# EPICS SNL sequencer program: injectorApp/src/injectorRampe_C2.stt
/*
#  C.E.A. IRFU/SIS/LDISC
#
#
#
*/
/*
*-----------------------------------------------------------------------
*   IFMIF/EVEDA Injecteur:
*   snl_Rampe_C2 : programme SNL pour la gestion de la commande de
*            rampe de COIL02_PS
*-----------------------------------------------------------------------
*/

/*program snl_Rampe_C2*/

program injectorRampe_C2

short OK_Rampe;
assign OK_Rampe to "SRC:COIL02_PS:PretRampe";
monitor OK_Rampe;

short Envoi_Rampe;
assign Envoi_Rampe to "SRC:COIL02_PS:RampeCmd";
monitor Envoi_Rampe;

ss ss1
{

        state connected {
             when ( (delay(2.0)) && (pvConnectCount() == pvChannelCount()) ) {
              printf("SNL_Rampe_C2 :entree programme - connexions etablies \n");

             } state Debut
       }

	state Debut
		   {
		      when ( (delay(1)) && ((OK_Rampe) == 1)) {
                         printf("ENVOI Start Rampe C2; \n");
                        Envoi_Rampe = 1;
                        pvPut(Envoi_Rampe);
                        OK_Rampe = 0;
                        pvPut(OK_Rampe);
                      } state suite_1
      }

	state suite_1
		{
	    	  when (delay(1)) {
                        printf("Fin sequence Envoi Start Rampe C2; \n");
                        Envoi_Rampe = 0;
                        pvPut(Envoi_Rampe);
                  } state Debut
     }
}
